(* IEC 61131-3 sources: SortJet_MasterSPS_Aufbau.fbsproj/08_POUs/Basis Funktionen, 41 files *)

(* ---- AuftragsdatenPruefen.fn.st ---- *)
(* METADATA
{
	"v3Meta": {
		"objectGuid": "657d7773-50f6-4a46-b86f-6fc5131c38e4"
	}
}
*)
FUNCTION AuftragsdatenPruefen : BOOL
VAR_INPUT

  // WORD
  wpMmiNummer  : WORD; // Stationsnummer von der die Auftraege geprueft werden sollen
  wpWandNr     : WORD; // Wandnummer von der die Auftraege geprueft werden sollen

  // STRUKT
  pData   : Auftragsdaten_ST;

END_VAR
VAR
  Basis : REFERENCE TO StationBasisParameter_ST;
END_VAR
Basis REF= getBasis(wpMmiNummer);
AuftragsdatenPruefen := TRUE;

// Glaslänge
IF ( pData.rAuftragsLaenge > Basis.stMKs.stGlasdaten[wpWandNr].rlMaxGlasLaenge ) THEN
  wpgFehlerdaten[0] := wpMmiNummer;
  wpgFehlerdaten[1] := REAL_TO_WORD(Basis.stMKs.stGlasdaten[wpWandNr].rlMaxGlasLaenge);
  wpgFehlerdaten[2] := REAL_TO_WORD(pData.rAuftragsLaenge);
  SpsError( eFehler_Station,
            cMELDUNG_AUFTRAGSDATEN_GLAS_ZU_LANG,
            wpMmiNummer,
            AutomatikkreisBestimmen(wpMmiNummer),
            wpgFehlerdaten );
  AuftragsdatenPruefen:=FALSE;
END_IF

IF ( pData.rAuftragsLaenge < Basis.stMKs.stGlasdaten[wpWandNr].rlMinGlasLaenge ) THEN
  wpgFehlerdaten[0] := wpMmiNummer;
  wpgFehlerdaten[1] := REAL_TO_WORD(Basis.stMKs.stGlasdaten[wpWandNr].rlMinGlasLaenge);
  wpgFehlerdaten[2] := REAL_TO_WORD(pData.rAuftragsLaenge);
  SpsError( eFehler_Station,
            cMELDUNG_AUFTRAGSDATEN_GLAS_ZU_KURZ,
            wpMmiNummer,
            AutomatikkreisBestimmen(wpMmiNummer),
            wpgFehlerdaten );
  AuftragsdatenPruefen:=FALSE;
END_IF

// Glashöhe
IF ( pData.rAuftragsHoehe > Basis.stMKs.stGlasdaten[wpWandNr].rlMaxGlasHoehe ) THEN
  wpgFehlerdaten[0] := wpMmiNummer;
  wpgFehlerdaten[1] := REAL_TO_WORD(Basis.stMKs.stGlasdaten[wpWandNr].rlMaxGlasHoehe);
  wpgFehlerdaten[2] := REAL_TO_WORD(pData.rAuftragsHoehe);
  SpsError( eFehler_Station,
            cMELDUNG_AUFTRAGSDATEN_GLAS_ZU_HOCH,
            wpMmiNummer,
            AutomatikkreisBestimmen(wpMmiNummer),
            wpgFehlerdaten );
  AuftragsdatenPruefen:=FALSE;
END_IF

IF ( pData.rAuftragsHoehe <  Basis.stMKs.stGlasdaten[wpWandNr].rlMinGlasHoehe ) THEN
  wpgFehlerdaten[0] := wpMmiNummer;
  wpgFehlerdaten[1] := REAL_TO_WORD(Basis.stMKs.stGlasdaten[wpWandNr].rlMinGlasHoehe);
  wpgFehlerdaten[2] := REAL_TO_WORD(pData.rAuftragsHoehe);
  SpsError( eFehler_Station,
            cMELDUNG_AUFTRAGSDATEN_GLAS_ZU_NIEDRIG,
            wpMmiNummer,
            AutomatikkreisBestimmen(wpMmiNummer),
            wpgFehlerdaten );
  AuftragsdatenPruefen:=FALSE;
END_IF

// Glasdicke
IF ( pData.rAuftragsDicke > Basis.stMKs.stGlasdaten[wpWandNr].rlMaxGlasDicke ) THEN
  wpgFehlerdaten[0] := wpMmiNummer;
  wpgFehlerdaten[1] := REAL_TO_WORD(Basis.stMKs.stGlasdaten[wpWandNr].rlMaxGlasDicke);
  wpgFehlerdaten[2] := REAL_TO_WORD(pData.rAuftragsDicke);
  SpsError( eFehler_Station,
            cMELDUNG_AUFTRAGSDATEN_GLAS_ZU_DICK,
            wpMmiNummer,
            AutomatikkreisBestimmen(wpMmiNummer),
            wpgFehlerdaten );
  AuftragsdatenPruefen := FALSE;
END_IF

IF ( pData.rAuftragsDicke < Basis.stMKs.stGlasdaten[wpWandNr].rlMinGlasDicke ) THEN
  wpgFehlerdaten[0] := wpMmiNummer;
  wpgFehlerdaten[1] := REAL_TO_WORD(Basis.stMKs.stGlasdaten[wpWandNr].rlMinGlasDicke);
  wpgFehlerdaten[2] := REAL_TO_WORD(pData.rAuftragsDicke);
  SpsError( eFehler_Station,
            cMELDUNG_AUFTRAGSDATEN_GLAS_ZU_DUENN,
            wpMmiNummer,
            AutomatikkreisBestimmen(wpMmiNummer),
            wpgFehlerdaten );
  AuftragsdatenPruefen := FALSE;
END_IF
END_FUNCTION

(* ---- AuftragsdatenUmkopieren.fn.st ---- *)
(* METADATA
{
	"v3Meta": {
		"objectGuid": "c0c5d446-5c0c-4964-91ed-f4edd34c4197"
	}
}
*)
FUNCTION AuftragsdatenUmkopieren : Auftragsdaten_ST
VAR_INPUT

  // BOOL
  bpAuswahlTransferstation_2  : BOOL := FALSE;
  bpAnwahlDurchtransport : BOOL := FALSE;

  // STRUCT
  stpAuftrag : Auftragsdaten_ST;

END_VAR
VAR

  // STRUCT
  stMerkerAuftrag  : Auftragsdaten_ST;

END_VAR
//-------------------------------------------------------------------------------------------------
// BAUSTEIN: LOGIK
//-------------------------------------------------------------------------------------------------

(* Hinweis:
   - Auftrag zwischenspeichern
*)
stMerkerAuftrag := stpAuftrag;

(* Hinweis:
   - Auftrag manipulieren
*)
IF ( NOT bpAuswahlTransferstation_2 AND NOT bpAnwahlDurchtransport ) THEN

  stMerkerAuftrag.wStationsNr            := stpAuftrag.wTransferstationsNr1;
  stMerkerAuftrag.wStationsWand          := stpAuftrag.wTransferwand;
  stMerkerAuftrag.rStationsZielposition  := stpAuftrag.rTransferposition1;
  stMerkerAuftrag.rVorabPosition         := stpAuftrag.rTransferposition1;

  stMerkerAuftrag.wTransferstationsNr1   := stpAuftrag.wStationsNr;
  stMerkerAuftrag.rTransferposition1     := stpAuftrag.rStationsZielposition;
  stMerkerAuftrag.wTransferwand          := stpAuftrag.wStationsWand;

ELSIF ( bpAnwahlDurchtransport ) THEN

  stMerkerAuftrag.wStationsNr            := stpAuftrag.wTransferstationsNr2;
  stMerkerAuftrag.wStationsWand          := stpAuftrag.wTransferwand;
  stMerkerAuftrag.rStationsZielposition  := stpAuftrag.rTransferposition2;
  stMerkerAuftrag.rVorabPosition         := stpAuftrag.rTransferposition2;

  stMerkerAuftrag.wTransferstationsNr2   := stpAuftrag.wStationsNr;
  stMerkerAuftrag.rTransferposition2     := stpAuftrag.rStationsZielposition;
  stMerkerAuftrag.wTransferwand          := stpAuftrag.wStationsWand;

ELSE
  stMerkerAuftrag.wStationsNr            := stpAuftrag.wTransferstationsNr2;
  stMerkerAuftrag.wStationsWand          := stpAuftrag.wTransferwand;
  stMerkerAuftrag.rStationsZielposition  := stpAuftrag.rTransferposition2;
  stMerkerAuftrag.rVorabPosition         := stpAuftrag.rTransferposition2;

  stMerkerAuftrag.wTransferstationsNr1   := stpAuftrag.wStationsNr;
  stMerkerAuftrag.rTransferposition1     := stpAuftrag.rStationsZielposition;
  stMerkerAuftrag.wTransferwand          := stpAuftrag.wStationsWand;

END_IF

AuftragsdatenUmkopieren := stMerkerAuftrag;
END_FUNCTION

(* ---- AutomatikAktiv.fn.st ---- *)
(* METADATA
{
	"v3Meta": {
		"objectGuid": "339b2ef9-3f23-482c-98f4-06c495d9a955"
	}
}
*)
FUNCTION AutomatikAktiv : BOOL
VAR_INPUT
  wpMmiNummer : WORD;
END_VAR
VAR
  wlIndex : WORD;
  Basis   : REFERENCE TO StationBasisParameter_ST;
END_VAR

// Hinweis:
// - Prueft ob einer der Automatikkreise der Station (Shuttle, TS, Station, Faecherwagen, Fremdanlage) aktiv ist
// - Die Basis wird ueber getBasis bestimmt
// - Unbekannte Nummer oder nicht zugewiesene MK => FALSE
// - Ein nicht belegter Automatikkreis (0) beendet die Pruefung
AutomatikAktiv := FALSE;

Basis REF= getBasis( wpMmiNummer );

IF NOT __ISVALIDREF( Basis ) THEN
  RETURN;
END_IF

IF NOT __ISVALIDREF( Basis.stMKs ) THEN
  RETURN;
END_IF

FOR wlIndex := cERSTER_AUTOMATIKKREIS TO cANZAHL_AUTOMATIKKREISE DO

  IF Basis.stMKs.eaAutomatikkreis[wlIndex] = 0 THEN
    RETURN;
  END_IF

  IF M_Automatik_Aktiv[Basis.stMKs.eaAutomatikkreis[wlIndex]] THEN
    AutomatikAktiv := TRUE;
    RETURN;
  END_IF

END_FOR
END_FUNCTION

(* ---- AutomatikFehlerSetzen.fn.st ---- *)
(* METADATA
{
	"v3Meta": {
		"objectGuid": "10c1b2d6-77ce-44d1-9dc1-390f3ff85d9b"
	}
}
*)
FUNCTION AutomatikFehlerSetzen : BOOL
VAR_INPUT
  eaAutomatikkreise : ARRAY[cERSTER_AUTOMATIKKREIS..cANZAHL_AUTOMATIKKREISE] OF Automatikkreis_EN;
  abpFehler : REFERENCE TO ARRAY[cERSTER_AUTOMATIKKREIS..cLETZTER_AUTOMATIKKREIS] OF BOOL;
END_VAR
VAR
  wlIndex: WORD;
END_VAR

FOR wlIndex := cERSTER_AUTOMATIKKREIS TO cANZAHL_AUTOMATIKKREISE DO

  IF eaAutomatikkreise[wlIndex] <> 0 THEN
    abpFehler[eaAutomatikkreise[wlIndex]] := TRUE;
  END_IF

END_FOR

AutomatikFehlerSetzen := TRUE;
END_FUNCTION

(* ---- AutomatikFehlerTransfershuttleSetzen.fn.st ---- *)
(* METADATA
{
	"v3Meta": {
		"objectGuid": "9a4c379e-af86-4c9e-b628-bbb819ee7aed"
	}
}
*)
FUNCTION AutomatikFehlerTransfershuttleSetzen : BOOL
VAR_INPUT
  eaAutomatikkreise    : ARRAY[cERSTER_AUTOMATIKKREIS..cANZAHL_AUTOMATIKKREISE] OF Automatikkreis_EN;
  abpFehler            : REFERENCE TO ARRAY[cERSTER_AUTOMATIKKREIS..cLETZTER_AUTOMATIKKREIS] OF BOOL;
  wSpeicherseiteFehler : BYTE; // cSPEICHER_EINLAUFSEITE oder cSPEICHER_AUSLAUFSEITE
END_VAR

// Hinweis:
// - Ein TS liegt meist als Trennglied unter dem Speicher in 2 AKs:
//   AK 1 = Einlaufseite, AK 2 = Auslaufseite
// - Welche Seite betroffen ist (Ein-/Austransport, rueckwaerts, Betriebsstopp)
//   entscheidet der Aufrufer in Job_Shuttle

// TS hat nur einen AK
IF ( eaAutomatikkreise[1] <> 0 AND eaAutomatikkreise[2] = 0 ) THEN
  abpFehler[eaAutomatikkreise[1]] := TRUE;

// TS hat 2 AK
ELSIF ( eaAutomatikkreise[1] <> 0 AND eaAutomatikkreise[2] <> 0 ) THEN
  IF ( wSpeicherseiteFehler = cSPEICHER_EINLAUFSEITE ) THEN
    abpFehler[eaAutomatikkreise[1]] := TRUE;
  ELSIF ( wSpeicherseiteFehler = cSPEICHER_AUSLAUFSEITE ) THEN
    abpFehler[eaAutomatikkreise[2]] := TRUE;
  END_IF
END_IF

AutomatikFehlerTransfershuttleSetzen := TRUE;
END_FUNCTION

(* ---- AutomatikkreisBestimmen.fn.st ---- *)
(* METADATA
{
	"v3Meta": {
		"objectGuid": "9ed7362d-6e8b-45fc-aaf5-a3cbb726335b"
	}
}
*)
FUNCTION AutomatikkreisBestimmen : Automatikkreis_EN
VAR_INPUT
  wpMmiNummer : WORD;
END_VAR
VAR
  Basis : REFERENCE TO StationBasisParameter_ST;
END_VAR

// Hinweis:
// - Erster Automatikkreis der Station (Shuttle, TS, Station, Faecherwagen, Fremdanlage) ueber getBasis
// - Unbekannte Nummer oder nicht zugewiesene MK => 0
AutomatikkreisBestimmen := 0;

Basis REF= getBasis( wpMmiNummer );

IF NOT __ISVALIDREF( Basis ) THEN
  RETURN;
END_IF

IF NOT __ISVALIDREF( Basis.stMKs ) THEN
  RETURN;
END_IF

AutomatikkreisBestimmen := Basis.stMKs.eaAutomatikkreis[cERSTER_AUTOMATIKKREIS];
END_FUNCTION

(* ---- BitToggleWord.fn.st ---- *)
(* METADATA
{
	"v3Meta": {
		"objectGuid": "aa0bc2f8-efb2-48a1-91f1-3637f8b86daf"
	}
}
*)
FUNCTION BitToggleWord : WORD
VAR_INPUT

  // WORD
  IN : WORD;

  // INT
  POS : INT;

END_VAR
//-------------------------------------------------------------------------------------------------
// BAUSTEIN: LOGIK
//-------------------------------------------------------------------------------------------------

(* Hinweis:
   - Diese Funktion setzt in einem WORD ein BIT an einer Position
     => Oscat-Lib
*)
BitToggleWord := SHL(WORD#1, POS) XOR IN;
END_FUNCTION

(* ---- checkSafetyCircuitAffectsComponent.fn.st ---- *)
(* METADATA
{
	"v3Meta": {
		"objectGuid": "b2891e00-4397-4c85-8733-7380e4011fc3"
	}
}
*)
FUNCTION checkSafetyCircuitAffectsComponent : BOOL
VAR_INPUT
  StationData  : REFERENCE TO StationBasisParameter_ST;
  SaftyCircuit : WORD;              // Sicherheitskreis
  eKomponente  : SK_Komponente_EN;  // Abgefragte Komponente (eSKKomponente_Alles = jeder SK zaehlt)
END_VAR
VAR
  wIndexMK : WORD := 0;
END_VAR
// Prueft, ob ein Sicherheitskreis die angegebene Komponente der Station abschaltet.
// - eSKKomponente_Alles: jeder SK der Station zaehlt -> TRUE
// - Standard (keine Teilabschaltung fuer diesen SK konfiguriert): SK schaltet alles ab -> TRUE
// - Mit Teilabschaltung: SK schaltet nur die markierten Komponenten ab

checkSafetyCircuitAffectsComponent := TRUE;

IF ( eKomponente = eSKKomponente_Alles ) THEN
  RETURN;
END_IF

FOR wIndexMK := 0 TO cANZAHL_SICHERHEITSKREISE DO
  IF     ( StationData.stMKs.astSicherheitskreisTeilabschaltung[wIndexMK].eSicherheitskreis = SaftyCircuit )
     AND StationData.stMKs.astSicherheitskreisTeilabschaltung[wIndexMK].bTeilabschaltung
  THEN
    CASE eKomponente OF
      eSKKomponente_Glastransport:   checkSafetyCircuitAffectsComponent := StationData.stMKs.astSicherheitskreisTeilabschaltung[wIndexMK].bGlastransport;
      eSKKomponente_Geblaese:        checkSafetyCircuitAffectsComponent := StationData.stMKs.astSicherheitskreisTeilabschaltung[wIndexMK].bGeblaese;
      eSKKomponente_Drehen:          checkSafetyCircuitAffectsComponent := StationData.stMKs.astSicherheitskreisTeilabschaltung[wIndexMK].bDrehen;
      eSKKomponente_Kippen:          checkSafetyCircuitAffectsComponent := StationData.stMKs.astSicherheitskreisTeilabschaltung[wIndexMK].bKippen;
      eSKKomponente_Querfahrt:       checkSafetyCircuitAffectsComponent := StationData.stMKs.astSicherheitskreisTeilabschaltung[wIndexMK].bQuerfahrt;
      eSKKomponente_Pneumatik:       checkSafetyCircuitAffectsComponent := StationData.stMKs.astSicherheitskreisTeilabschaltung[wIndexMK].bPneumatik;
      eSKKomponente_Greifer:         checkSafetyCircuitAffectsComponent := StationData.stMKs.astSicherheitskreisTeilabschaltung[wIndexMK].bGreifer;
      eSKKomponente_Wandverstellung: checkSafetyCircuitAffectsComponent := StationData.stMKs.astSicherheitskreisTeilabschaltung[wIndexMK].bWandverstellung;
      eSKKomponente_Messachse:       checkSafetyCircuitAffectsComponent := StationData.stMKs.astSicherheitskreisTeilabschaltung[wIndexMK].bMessachse;
    END_CASE
    RETURN;
  END_IF
END_FOR
END_FUNCTION

(* ---- checkSafetyCircuits.fn.st ---- *)
(* METADATA
{
	"v3Meta": {
		"objectGuid": "a5602391-f145-45a7-88a7-cf2977d4c874"
	}
}
*)
FUNCTION checkSafetyCircuits : BOOL
VAR_INPUT
  StationData  : REFERENCE TO StationBasisParameter_ST;
  SaftyCircuit : WORD;
END_VAR
VAR
  wIndexMK : WORD := 0;
END_VAR
// It will checked if the safety circuit configured for this station

checkSafetyCircuits := FALSE;

FOR wIndexMK := 0 TO cANZAHL_SICHERHEITSKREISE DO
  IF ( SaftyCircuit = StationData.stMKs.eaSicherheitskreis[wIndexMK] ) THEN
    checkSafetyCircuits := TRUE;
    EXIT;
  END_IF
END_FOR
END_FUNCTION

(* ---- checkSafetyCircuitsClosed.fn.st ---- *)
(* METADATA
{
	"v3Meta": {
		"objectGuid": "1a45708a-46ce-48f5-a3b2-b0c20261c8e1"
	}
}
*)
FUNCTION checkSafetyCircuitsClosed : BOOL
VAR_INPUT
  StationData : REFERENCE TO StationBasisParameter_ST;
  eKomponente : SK_Komponente_EN := eSKKomponente_Alles; // Optional: Pruefung fuer eine Komponente (beruecksichtigt Teilabschaltung), Standard: jeder SK zaehlt
END_VAR
VAR
  arrCircuits : ARRAY[cERSTER_SICHERHEITSKREIS..cLETZTER_SICHERHEITSKREIS] OF BOOL;
  wIndex   : WORD := 0;
  wIndexMK : WORD := 0;
END_VAR
// It will checked if the safety circuit is activ

checkSafetyCircuitsClosed := TRUE;

FOR wIndex := cERSTER_SICHERHEITSKREIS TO cLETZTER_SICHERHEITSKREIS DO
  arrCircuits[wIndex] := Sicherheitskreis[wIndex].bpSicherheitskreisGeschlossen;
END_FOR

FOR wIndex := cERSTER_SICHERHEITSKREIS TO cLETZTER_SICHERHEITSKREIS DO
  FOR wIndexMK := 0 TO cANZAHL_SICHERHEITSKREISE DO
    IF ( wIndex = StationData.stMKs.eaSicherheitskreis[wIndexMK] ) THEN
      IF NOT arrCircuits[wIndex] AND checkSafetyCircuitAffectsComponent(StationData, wIndex, eKomponente) THEN
        checkSafetyCircuitsClosed := FALSE;
      END_IF
    END_IF
  END_FOR
END_FOR
END_FUNCTION

(* ---- checkSafetyCircuitsClosedFromAutomaticCircuit.fn.st ---- *)
(* METADATA
{
	"v3Meta": {
		"objectGuid": "6a4b769b-603d-4996-8e76-e26c1b994362"
	}
}
*)
FUNCTION checkSafetyCircuitsClosedFromAutomaticCircuit : BOOL
VAR_INPUT

  // WORD
  wlAutomatikkreis : WORD;

  // BOOL
  bNurStartBlockierende : BOOL := FALSE; // TRUE: nur Sicherheitskreise beruecksichtigen, die Systemcheck und Initialisierung blockieren [MK bBlockiertStart]

END_VAR
VAR
  // BOOL
  findInWORDArray               : BOOL;
  bSicherheitskreisIstDurchgang : BOOL;

  // WORD
  wlIndexSicherheitskreis : WORD;

  // ENUM
  INDEX : Automatikkreis_EN;

END_VAR

// DIESE FUNKTION BERÜCKSICHTIGT KEINE DURCHGÄNGE !!!
checkSafetyCircuitsClosedFromAutomaticCircuit := TRUE;

FOR wlIndexSicherheitskreis := cERSTER_SICHERHEITSKREIS TO cLETZTER_SICHERHEITSKREIS DO

  bSicherheitskreisIstDurchgang := FALSE;

  FOR INDEX := cERSTER_DURCHGANG TO cANZAHL_DURCHGANGE DO
    IF apgMKDurchgang[INDEX].eZuBlockierenderSK = wlIndexSicherheitskreis THEN
      bSicherheitskreisIstDurchgang := TRUE;
      EXIT;
    END_IF
  END_FOR

  IF NOT bSicherheitskreisIstDurchgang THEN

    findInWORDArray := FALSE;

    FOR INDEX := cERSTER_AUTOMATIKKREIS TO cLETZTER_AUTOMATIKKREIS DO
      IF apgMKSicherheiskreis[wlIndexSicherheitskreis].eaAutomatikkreis[INDEX] = wlAutomatikkreis THEN
        findInWORDArray := TRUE;
        EXIT;
      END_IF
    END_FOR

    IF findInWORDArray AND ( NOT bNurStartBlockierende OR apgMKSicherheiskreis[wlIndexSicherheitskreis].bBlockiertStart ) THEN
      checkSafetyCircuitsClosedFromAutomaticCircuit :=
                                                      checkSafetyCircuitsClosedFromAutomaticCircuit
                                                      AND Sicherheitskreis[wlIndexSicherheitskreis].bpSicherheitskreisGeschlossen;
    END_IF

  END_IF

END_FOR
END_FUNCTION

(* ---- checkSafetyCircuitsConfigured.fn.st ---- *)
(* METADATA
{
	"v3Meta": {
		"objectGuid": "dcded4cc-d766-4c84-a212-2fe6cc93f6db"
	}
}
*)
FUNCTION checkSafetyCircuitsConfigured : BOOL
VAR_INPUT
  StationData : REFERENCE TO StationBasisParameter_ST;
END_VAR
VAR
  wIndexMK : WORD := 0;
END_VAR

// It will checked if a safety circuit is configured

checkSafetyCircuitsConfigured := FALSE;

IF NOT __ISVALIDREF(StationData.stMKs) OR_ELSE StationData.stMKs.bDeaktivieren THEN
  RETURN;
END_IF

FOR wIndexMK := 0 TO cANZAHL_SICHERHEITSKREISE DO
  IF ( StationData.stMKs.eaSicherheitskreis[wIndexMK] <> eSicherheitskreis_Undefiniert ) THEN
    checkSafetyCircuitsConfigured := TRUE;
    EXIT;
  END_IF
END_FOR
END_FUNCTION

(* ---- checkSafetyCircuitsNotBlocked.fn.st ---- *)
(* METADATA
{
	"v3Meta": {
		"objectGuid": "93537a12-23ea-4a31-94f7-53154eb0b75f"
	}
}
*)
FUNCTION checkSafetyCircuitsNotBlocked : BOOL
VAR_INPUT
  StationData : REFERENCE TO StationBasisParameter_ST;
  eKomponente : SK_Komponente_EN := eSKKomponente_Alles; // Optional: Pruefung fuer eine Komponente (beruecksichtigt Teilabschaltung), Standard: jeder SK zaehlt
END_VAR
VAR
  arrCircuits : ARRAY[cERSTER_SICHERHEITSKREIS..cLETZTER_SICHERHEITSKREIS] OF BOOL;
  wIndex   : WORD := 0;
  wIndexMK : WORD := 0;
END_VAR
// It will checked if the safety circuit is activ

checkSafetyCircuitsNotBlocked := TRUE;

FOR wIndex := cERSTER_SICHERHEITSKREIS TO cLETZTER_SICHERHEITSKREIS DO
  arrCircuits[wIndex] :=         Sicherheitskreis[wIndex].bpSicherheitskreisGeschlossen
                                 AND NOT Sicherheitskreis[wIndex].bpStationenBlocken
                                 AND NOT Sicherheitskreis[wIndex].bpAnforderungSKGestellt
                                 AND NOT Sicherheitskreis[wIndex].bpAnforderungSicherheitkreisAusloesen;
END_FOR

FOR wIndex := cERSTER_SICHERHEITSKREIS TO cLETZTER_SICHERHEITSKREIS DO
  FOR wIndexMK := 0 TO cANZAHL_SICHERHEITSKREISE DO
    IF ( wIndex = StationData.stMKs.eaSicherheitskreis[wIndexMK] ) THEN
      IF ( ( NOT arrCircuits[wIndex] ) AND ( NOT bgSicherheitstechnikBruecken ) AND checkSafetyCircuitAffectsComponent(StationData, wIndex, eKomponente) ) THEN
        checkSafetyCircuitsNotBlocked := FALSE;
        EXIT;
      END_IF
    END_IF
  END_FOR
END_FOR
END_FUNCTION

(* ---- checkSafetyCircuitsRequested.fn.st ---- *)
(* METADATA
{
	"v3Meta": {
		"objectGuid": "c6e29fd6-ba36-47ef-8c35-03485548b8fc"
	}
}
*)
FUNCTION checkSafetyCircuitsRequested : BOOL
VAR_INPUT
  StationData : REFERENCE TO StationBasisParameter_ST;
  eKomponente : SK_Komponente_EN := eSKKomponente_Alles; // Optional: Pruefung fuer eine Komponente (beruecksichtigt Teilabschaltung), Standard: jeder SK zaehlt
END_VAR
VAR
  arrCircuits : ARRAY[cERSTER_SICHERHEITSKREIS..cLETZTER_SICHERHEITSKREIS] OF BOOL;
  wIndex   : WORD := 0;
  wIndexMK : WORD := 0;
END_VAR
// It will checked if the safety circuit is requested

checkSafetyCircuitsRequested := TRUE;

FOR wIndex := cERSTER_SICHERHEITSKREIS TO cLETZTER_SICHERHEITSKREIS DO
  arrCircuits[wIndex] :=         Sicherheitskreis[wIndex].bpSicherheitskreisGeschlossen
                                 AND NOT Sicherheitskreis[wIndex].bpAnforderungSKGestellt;
END_FOR

FOR wIndex := cERSTER_SICHERHEITSKREIS TO cLETZTER_SICHERHEITSKREIS DO

  FOR wIndexMK := 0 TO cANZAHL_SICHERHEITSKREISE DO
    IF ( wIndex = StationData.stMKs.eaSicherheitskreis[wIndexMK] ) THEN
      IF NOT arrCircuits[wIndex] AND checkSafetyCircuitAffectsComponent(StationData, wIndex, eKomponente) THEN
        checkSafetyCircuitsRequested := FALSE;
      END_IF
    END_IF
  END_FOR
END_FOR
END_FUNCTION

(* ---- DEC.fn.st ---- *)
(* METADATA
{
	"v3Meta": {
		"objectGuid": "e4081493-5d9a-4e63-8c4b-cba513ba3d02"
	}
}
*)
{attribute 'excludefrombuild'}
FUNCTION DEC : INT
VAR_INPUT
  iWert    : INT;
  iMinuend : INT;
END_VAR

(* Hinweis:
   - Funktion zum reduzieren der Eingangsvariablen X um 1.
*)
DEC := iWert - iMinuend;
END_FUNCTION

(* ---- findInWORDArray.fn.st ---- *)
(* METADATA
{
	"v3Meta": {
		"objectGuid": "27266190-4c13-454c-9114-87648310c4ec"
	}
}
*)
FUNCTION findInWORDArray : BOOL
VAR_INPUT
  awpArray : ARRAY[1..10] OF WORD;
  wpValueToFind : WORD;
END_VAR
VAR
  INDEX : WORD;
END_VAR

findInWORDArray := FALSE;

FOR INDEX := 1 TO 10 DO

  IF awpArray[INDEX] = wpValueToFind THEN
    findInWORDArray := TRUE;
    EXIT;
  END_IF

END_FOR
END_FUNCTION

(* ---- getAnzahlSystemcheckZyklen.fn.st ---- *)
(* METADATA
{
	"v3Meta": {
		"objectGuid": "64956d77-da35-4a2e-90f0-c969659e6e9b"
	}
}
*)
FUNCTION getAnzahlSystemcheckZyklen : WORD
VAR_INPUT
END_VAR
VAR
  wIndex : WORD;
  bByte  : BYTE;
  ptNull : REFERENCE TO BYTE := 0;
END_VAR

getAnzahlSystemcheckZyklen := 0;

// Alle Shuttles durchlaufen
FOR wIndex := cERSTES_SHUTTLE TO cLETZTES_SHUTTLE DO
  // Null-Pointer wenn kein Zyklus in den MKs zugewiesen wurde
  IF starrShuttleBasisParameter[wIndex].stMKs.eSystemcheckZyklus = eSystemcheckZyklus_Undefiniert THEN
    SysExceptGenerateException( RtsExceptions.RTSEXCPT_ARRAYBOUNDS );
  //bByte := ptNull; (*cause access violation *)
  ELSE // Ansonsten den definierten Zyklus in das Array übernehmen
    // Neuer höherer Wert? Dann wegspeichern
    IF getAnzahlSystemcheckZyklen < starrShuttleBasisParameter[wIndex].stMKs.eSystemcheckZyklus THEN
      getAnzahlSystemcheckZyklen := starrShuttleBasisParameter[wIndex].stMKs.eSystemcheckZyklus;
    END_IF
  END_IF
END_FOR

// Alle Stationen durchlaufen
FOR wIndex := cERSTE_STATION TO cLETZTE_STATION DO
  // Null-Pointer wenn kein Zyklus in den MKs zugewiesen wurde
  IF NOT __ISVALIDREF(starrStationBasisParameter[wIndex].stMKs) THEN
    CONTINUE;
  ELSIF starrStationBasisParameter[wIndex].stMKs.eSystemcheckZyklus = eSystemcheckZyklus_Undefiniert AND NOT starrStationBasisParameter[wIndex].stMKs.bDeaktivieren THEN
    SysExceptGenerateException( RtsExceptions.RTSEXCPT_ARRAYBOUNDS );
  //bByte := ptNull; (*cause access violation *)
  ELSE // Ansonsten den definierten Zyklus in das Array übernehmen
    // Neuer höherer Wert? Dann wegspeichern
    IF getAnzahlSystemcheckZyklen < starrStationBasisParameter[wIndex].stMKs.eSystemcheckZyklus THEN
      getAnzahlSystemcheckZyklen := starrStationBasisParameter[wIndex].stMKs.eSystemcheckZyklus;
    END_IF
  END_IF
END_FOR

// Null-Pointer wenn kein Ergebnis gefunden wurde (fehlerhafter Zustand)
IF ( getAnzahlSystemcheckZyklen = 0 ) THEN
  SysExceptGenerateException( RtsExceptions.RTSEXCPT_ARRAYBOUNDS );
//bByte := ptNull; (*cause access violation *)
END_IF
END_FUNCTION

(* ---- getAuftragsdaten.fn.st ---- *)
(* METADATA
{
	"v3Meta": {
		"objectGuid": "e09c3e56-23fc-432f-9a18-960dccfa6275"
	}
}
*)
FUNCTION getAuftragsdaten : REFERENCE TO Auftragsdaten_ST
VAR_INPUT

  // WORD
  wpMmiNummer  : WORD; // Stationsnummer, deren aktueller Auftrag geliefert werden soll
  wpWand       : WORD; // Wand (nur Shuttles und Stationen)

END_VAR
// Hinweis:
// - Gegenstueck zu getBasis: liefert den aktuellen Job-Auftrag einer Station
// - Ungueltige Nummer oder Wand => ungueltige Referenz (Aufrufer prueft mit __ISVALIDREF)
CASE wpMmiNummer OF

  cERSTES_SHUTTLE..cLETZTES_SHUTTLE:
    IF ( PruefungWertImIntervall( wpWand, cWAND_1, cANZAHL_WAENDE ) ) THEN
      getAuftragsdaten REF= Job_Shuttle.AuftragsdatenWand[wpMmiNummer, wpWand];
    END_IF

  cERSTES_TRANSFERSHUTTLE..cLETZTES_TRANSFERSHUTTLE:
    getAuftragsdaten REF= Job_Shuttle.AuftragsdatenTransfershuttle[wpMmiNummer];

  cERSTE_STATION..cLETZTE_STATION:
    IF ( PruefungWertImIntervall( wpWand, cWAND_1, cANZAHL_WAENDE ) ) THEN
      getAuftragsdaten REF= Job_Stationen.AuftragsdatenWand[wpMmiNummer, wpWand];
    END_IF

  cERSTE_FREMDANLAGE_AUSLAUF..cLETZTE_FREMDANLAGE_EINLAUF:
    getAuftragsdaten REF= Job_Fremdanlage.AuftragsdatenFremdanlage[wpMmiNummer];

END_CASE
END_FUNCTION

(* ---- getBasis.fn.st ---- *)
(* METADATA
{
	"v3Meta": {
		"objectGuid": "cb0abf05-d74d-4b59-9143-e94abaf551fa"
	}
}
*)
FUNCTION getBasis : REFERENCE TO  StationBasisParameter_ST
VAR_INPUT

  // WORD
  wpMmiNummer  : WORD; // Stationsnummer von der die Auftraege geprueft werden sollen

END_VAR
CASE wpMmiNummer OF

  cERSTES_SHUTTLE..cLETZTES_SHUTTLE:
    getBasis REF= starrShuttleBasisParameter[wpMmiNummer];

  cERSTES_TRANSFERSHUTTLE..cLETZTES_TRANSFERSHUTTLE:
    getBasis REF= starrTransfershuttleBasisParameter[wpMmiNummer];

  cERSTE_STATION..cLETZTE_STATION:
    getBasis REF= starrStationBasisParameter[wpMmiNummer];

  cERSTE_FAECHERWAGENSTATIONS_NR..cLETZTE_FAECHERWAGENSTATIONS_NR:
    getBasis REF= starrFaecherwagenBasisParameter[wpMmiNummer];

  cERSTE_FREMDANLAGE_EINLAUF..cLETZTE_FREMDANLAGE_EINLAUF:
    getBasis REF= starrFremdanlageEinlaufStationBasisParameter[wpMmiNummer];

  cERSTE_FREMDANLAGE_AUSLAUF..cLETZTE_FREMDANLAGE_AUSLAUF:
    getBasis REF= starrFremdanlageAuslaufStationBasisParameter[wpMmiNummer];

END_CASE
END_FUNCTION

(* ---- GetBitFromWord.fn.st ---- *)
(* METADATA
{
	"v3Meta": {
		"objectGuid": "4ac38ee7-2639-4587-9c58-5882c3701cd8"
	}
}
*)
FUNCTION GetBitFromWord : Bool
VAR_INPUT
  Value : WORD;   // Das Wort, aus dem du die Bits auslesen willst
  Index : Word;    // Welches Bit (0..15)
END_VAR
VAR
END_VAR

GetBitFromWord := (Value AND SHL(1, Index)) <> 0;
END_FUNCTION

(* ---- getRealShuttleMaxPos.fn.st ---- *)
(* METADATA
{
	"v3Meta": {
		"objectGuid": "fdbd0502-3da4-4780-aa1a-b043617e0f01"
	}
}
*)
FUNCTION getRealShuttleMaxPos : REAL
VAR_INPUT
  wShuttleNummer : WORD;
END_VAR

getRealShuttleMaxPos := aShuttle[wShuttleNummer].Querfahrt.Antrieb.rpMaxPosition;
END_FUNCTION

(* ---- getRealShuttleMinPos.fn.st ---- *)
(* METADATA
{
	"v3Meta": {
		"objectGuid": "77446a83-5414-4511-a85e-8d0f27ae2e7b"
	}
}
*)
FUNCTION getRealShuttleMinPos : REAL
VAR_INPUT
  wShuttleNummer : WORD;
END_VAR

getRealShuttleMinPos := aShuttle[wShuttleNummer].Querfahrt.Antrieb.rpMinPosition;
END_FUNCTION

(* ---- GlasGewichtErmitteln.fn.st ---- *)
(* METADATA
{
	"v3Meta": {
		"objectGuid": "bd924e48-93d5-4f05-bff1-59051efc4e7c"
	}
}
*)
FUNCTION GlasGewichtErmitteln : REAL
VAR_INPUT

  // REAL
  rpGlaslaenge  : REAL := REAL#0; // [mm] -> Wert in mm
  rpGlasbreite  : REAL := REAL#0; // [mm] -> Wert in mm
  rpGlasstaerke : REAL := REAL#0; // [mm] -> Wert in mm

END_VAR
VAR

  // REAL
  rlErgebnis : REAL := REAL#0;
  rlLaenge   : REAL := REAL#0; // [mm] -> Wert in dm [UMRECHNUNG]
  rlBreite   : REAL := REAL#0; // [mm] -> Wert in dm [UMRECHNUNG]
  rlStaerke  : REAL := REAL#0; // [mm] -> Wert in dm [UMRECHNUNG]

END_VAR

VAR CONSTANT

  // WORD
  cUMRECHNUNG_MM_IN_DM      : REAL := 100.0;

  // REAL
  cSPEZIFISCHES_GLASGEWICHT : REAL := REAL#2.5; //IN kg/dm³

END_VAR

rlErgebnis := REAL#0;

rlLaenge  := rpGlaslaenge / cUMRECHNUNG_MM_IN_DM;
rlBreite  := rpGlasbreite / cUMRECHNUNG_MM_IN_DM;
rlStaerke := rpGlasstaerke/ cUMRECHNUNG_MM_IN_DM;

GlasGewichtErmitteln := ( ( rlLaenge * rlBreite * rlStaerke ) ) * cSPEZIFISCHES_GLASGEWICHT;
END_FUNCTION

(* ---- INC_UI.fn.st ---- *)
(* METADATA
{
	"v3Meta": {
		"objectGuid": "e071f047-ba29-40c0-bdd3-dce3563eb13b"
	}
}
*)
FUNCTION INC_UI : UINT
VAR_INPUT
  pui : REFERENCE TO UINT;
END_VAR
VAR
END_VAR

IF pui < 65536
THEN
  pui := pui + 1;
END_IF
END_FUNCTION

(* ---- INCI.fn.st ---- *)
(* METADATA
{
	"v3Meta": {
		"objectGuid": "47a21df2-edbb-49b0-932f-ef927933ed32"
	}
}
*)
FUNCTION INCI : INT
VAR_INPUT
  X : INT;
  N : INT;
END_VAR

(* Hinweis:
   - Funktion zum erhoehen der Eingangsvariablen X um 1. Sobald X den Wert N erreicht hat startet der Wert wieder bei 0.
*)
IF ( X >= N - 1 ) THEN
  INCI := 0;
ELSE
  INCI := X + 1;
END_IF;
END_FUNCTION

(* ---- INCW.fn.st ---- *)
(* METADATA
{
	"v3Meta": {
		"objectGuid": "c3800ee6-fccf-491b-bd53-b6c1155883a9"
	}
}
*)
FUNCTION INCW : WORD
VAR_INPUT
  X : WORD;
  N : WORD;
END_VAR

(* Hinweis:
   - Funktion zum erhoehen der Eingangsvariablen X um 1. Sobald X den Wert N erreicht hat startet der Wert wieder bei 0.
*)
IF ( X >= N - 1 ) THEN
  INCW := 0;
ELSE
  INCW := X + 1;
END_IF;
END_FUNCTION

(* ---- IsBetweenLReal.fn.st ---- *)
(* METADATA
{
	"v3Meta": {
		"objectGuid": "605f94de-cd86-43d0-95cd-83c44bc0f8dc"
	}
}
*)
FUNCTION IsBetweenLReal : BOOL
VAR_INPUT
  lriValue   : LREAL;
  lriBorder1 : LREAL;
  lriBorder2 : LREAL;
END_VAR
VAR
END_VAR

IsBetweenLReal := FALSE;

IF lriBorder1 < lriBorder2 THEN
  IsBetweenLReal := lriBorder1 <= lriValue
                    AND lriValue <= lriBorder2;
ELSE
  IsBetweenLReal := lriBorder2 <= lriValue
                    AND lriValue <= lriBorder1;
END_IF
END_FUNCTION

(* ---- IsBetweenWORD.fn.st ---- *)
(* METADATA
{
	"v3Meta": {
		"objectGuid": "640e1550-054d-48b5-a8dc-d9ce3f68325e"
	}
}
*)
FUNCTION IsBetweenWORD : BOOL
VAR_INPUT
  lwValue   : WORD;
  lwBorder1 : WORD;
  lwBorder2 : WORD;
END_VAR
VAR
END_VAR

IsBetweenWORD := FALSE;

IF lwBorder1 < lwBorder2 THEN
  IsBetweenWORD := lwBorder1 <= lwValue
                   AND lwValue <= lwBorder2;
ELSE
  IsBetweenWORD := lwBorder2 <= lwValue
                   AND lwValue <= lwBorder1;
END_IF
END_FUNCTION

(* ---- IsInRange.fn.st ---- *)
(* METADATA
{
	"v3Meta": {
		"objectGuid": "666a809c-7e52-4abd-9f01-34086fac7ebd"
	}
}
*)
FUNCTION IsInRange : BOOL
VAR_INPUT
  rlValue : REAL;
  rlTargetValue : REAL;
  rlThresshold : REAL;
END_VAR
VAR
END_VAR

IsInRange := ABS(rlValue - rlTargetValue) <= rlThresshold;
END_FUNCTION

(* ---- PruefungWertImIntervall.fn.st ---- *)
(* METADATA
{
	"v3Meta": {
		"objectGuid": "b7be4780-1c3e-4371-bb2a-cc9122a11be5"
	}
}
*)
FUNCTION PruefungWertImIntervall : BOOL
VAR_INPUT

  // WORD
  wpWert         : WORD;
  wpIntervallMin : WORD;
  wpIntervallMax : WORD;

END_VAR
VAR
END_VAR
//-------------------------------------------------------------------------------------------------
// LOGIK
//-------------------------------------------------------------------------------------------------
IF (  wpWert >= wpIntervallMin
     AND wpWert <= wpIntervallMax )
THEN
  PruefungWertImIntervall := TRUE;
ELSE
  PruefungWertImIntervall := FALSE;
END_IF
END_FUNCTION

(* ---- PruefungWertImIntervallAutomatikkreise.fn.st ---- *)
(* METADATA
{
	"v3Meta": {
		"objectGuid": "4fd29558-d6eb-46af-8028-798423b786a8"
	}
}
*)
FUNCTION PruefungWertImIntervallAutomatikkreise : BOOL
VAR_INPUT

  // WORD
  wpWert         : ARRAY[cERSTER_AUTOMATIKKREIS..cANZAHL_AUTOMATIKKREISE] OF Automatikkreis_EN;
  wpIntervallMin : WORD;
  wpIntervallMax : WORD;

END_VAR
VAR
  wlIndex : WORD;
END_VAR
//-------------------------------------------------------------------------------------------------
// LOGIK
//-------------------------------------------------------------------------------------------------
PruefungWertImIntervallAutomatikkreise := FALSE;

FOR wlIndex := cERSTER_AUTOMATIKKREIS TO cANZAHL_AUTOMATIKKREISE DO

  IF wpWert[wlIndex] = 0 THEN
    RETURN;
  END_IF

  IF (  wpWert[wlIndex] >= wpIntervallMin
       AND wpWert[wlIndex] <= wpIntervallMax )
  THEN
    PruefungWertImIntervallAutomatikkreise := TRUE;
  ELSE
    PruefungWertImIntervallAutomatikkreise := FALSE;
    RETURN;
  END_IF

END_FOR
END_FUNCTION

(* ---- RemoveETX.fn.st ---- *)
(* METADATA
{
	"v3Meta": {
		"objectGuid": "6a30dc93-6cfb-42ec-8e94-53fcaf08507e"
	}
}
*)
FUNCTION RemoveETX : ARRAY [0..3] OF DWORD
VAR_INPUT
  SheetID : ARRAY [0..3] OF DWORD;
END_VAR
VAR
  i, dwIn, dwOut, sh : INT;
  b : BYTE;
  tmp : DWORD;
END_VAR
FOR i := 0 TO 3 DO RemoveETX[i] := DWORD#0; END_FOR;

FOR i := 0 TO 15 DO
  dwIn := i / 4; sh := (i MOD 4) * 8;

  tmp := SHR(SheetID[dwIn], sh);     // byte runter schieben
  tmp := tmp MOD DWORD#256;          // entspricht AND 16#FF
  b := DWORD_TO_BYTE(tmp);

  IF b = BYTE#16#03 THEN b := BYTE#0; END_IF;

  dwOut := i / 4; sh := (i MOD 4) * 8;
  RemoveETX[dwOut] := RemoveETX[dwOut] + SHL(BYTE_TO_DWORD(b), sh);  // + statt OR
END_FOR;
END_FUNCTION

(* ---- ScheibenQuittierung.fn.st ---- *)
(* METADATA
{
	"v3Meta": {
		"objectGuid": "e5781056-5434-4b12-a4a2-e1c1e4aeb816"
	}
}
*)
FUNCTION ScheibenQuittierung : BOOL
VAR_INPUT

  // WORD
  wpQuellstation : WORD;
  wpZielStation  : WORD;
  wpQuellwand    : WORD := 1;
  wpZielwand     : WORD := 1;
  wpAuftragsTyp  : WORD := 0;

  // DWORD
  dwpWartezeit   : DWORD := 0;

END_VAR

VAR

  // BOOLEAN
  blResult : BOOL := FALSE;

END_VAR
//-------------------------------------------------------------------------------------------------
// FUNKTION: QUITTIEREN DER SCHEIBE
//-------------------------------------------------------------------------------------------------

wSps2MmiZielStation  := wpZielStation;
wSps2MmiQuellStation := wpQuellstation;
wSps2MmiZielWand     := wpZielwand;
wSps2MmiQuellWand    := wpQuellwand;
dwSps2MmiWartezeit   := dwpWartezeit;
wSPS2MMIAuftragstyp  := wpAuftragsTyp;

MsgToMmi(auftragsnr_w := SB0_SPS_QUIT_SHEET_ORDER );

ScheibenQuittierung := TRUE;
END_FUNCTION

(* ---- SendShuttlePosition.fn.st ---- *)
(* METADATA
{
	"v3Meta": {
		"objectGuid": "61256a4f-f80b-4fab-9669-5735e5c0be34"
	}
}
*)
FUNCTION SendShuttlePosition : BOOL
VAR_INPUT
END_VAR
VAR
  wlNummer : WORD;
  wlSlot   : WORD;
END_VAR
VAR CONSTANT
  cANZAHL_SLOTS_TELEGRAMM : WORD := 12; // Positionen die SB0_SPS_SORTIERUNGSHUTTLEPOS transportiert
END_VAR

//########################################## Changelog ################################################
//
//  2017-11-26 KV - Erstellt
//     => Function to send the current actual position of shuttle
//
//########################################## Changelog ################################################

(* Hinweis:
   - Die Position steht im MMI-Telegramm an einer festen Stelle (Slot), die Reihenfolge ist fest:
     1. Shuttles, 2. Transfershuttles, 3. Stationen die ein Shuttle sind [bStationIstShuttle]
   - Jede MK belegt einen Slot, auch wenn sie deaktiviert ist
   - Was nicht mehr ins Telegramm passt, wird nicht gesendet
*)
FOR wlSlot := 0 TO cANZAHL_SLOTS_TELEGRAMM - 1 DO
  rSps2MmiShuttlePosition[wlSlot] := 0.0;
END_FOR

wlSlot := 0;

// SHUTTLE
FOR wlNummer := cERSTES_SHUTTLE TO cLETZTES_SHUTTLE DO
  IF wlSlot < cANZAHL_SLOTS_TELEGRAMM THEN
    rSps2MmiShuttlePosition[wlSlot] := starrShuttleBasisParameter[wlNummer].rAktuellePositionQuerfahrt;
    wlSlot := wlSlot + 1;
  END_IF
END_FOR

// TRANSFERSHUTTLE
FOR wlNummer := cERSTES_TRANSFERSHUTTLE TO cLETZTES_TRANSFERSHUTTLE DO
  IF wlSlot < cANZAHL_SLOTS_TELEGRAMM THEN
    rSps2MmiShuttlePosition[wlSlot] := starrTransferShuttleBasisParameter[wlNummer].rAktuellePositionQuerfahrt;
    wlSlot := wlSlot + 1;
  END_IF
END_FOR

// STATIONEN die ein Shuttle sind
FOR wlNummer := cERSTE_STATION TO cLETZTE_STATION DO
  IF starrStationBasisParameter[wlNummer].stMKs.stSchnittstellendaten.bStationIstShuttle THEN
    IF wlSlot < cANZAHL_SLOTS_TELEGRAMM THEN
      rSps2MmiShuttlePosition[wlSlot] := starrStationBasisParameter[wlNummer].rAktuellePositionQuerfahrt;
      wlSlot := wlSlot + 1;
    END_IF
  END_IF
END_FOR

MsgToMmi(auftragsnr_w := SB0_SPS_SORTIERUNGSHUTTLEPOS);

SendShuttlePosition := TRUE;
END_FUNCTION

(* ---- setFreigabeKomponenten.fn.st ---- *)
(* METADATA
{
	"v3Meta": {
		"objectGuid": "691bf0f6-0a88-4d0a-9736-fcf4e429c02d"
	}
}
*)
FUNCTION setFreigabeKomponenten : BOOL
VAR_INPUT
  StationData : REFERENCE TO StationBasisParameter_ST;
END_VAR
VAR
  blSKAuswerten : BOOL; // Station hat gueltige MK, ist aktiv und hat mindestens einen SK konfiguriert
END_VAR
// Setzt alle Freigaben der Station (stFreigabe):
// - bAlles: NotHalt OK und ALLE Sicherheitskreise der Station geschlossen
// - bX    : NotHalt OK und alle SKs geschlossen, die Komponente X abschalten
//           (SK ohne Teilabschaltung schaltet alles ab, SK mit Teilabschaltung nur die markierten Komponenten)
// - Ohne konfigurierten SK (oder Station deaktiviert / keine MK): nur NotHalt
// - bgSicherheitstechnikBruecken setzt alle Freigaben

blSKAuswerten := checkSafetyCircuitsConfigured(StationData);

StationData.stFreigabe.bAlles           := ( NotHalt.bpNotHaltOK AND ( NOT blSKAuswerten OR_ELSE checkSafetyCircuitsClosed(StationData, eSKKomponente_Alles) ) )           OR bgSicherheitstechnikBruecken;
StationData.stFreigabe.bGlastransport   := ( NotHalt.bpNotHaltOK AND ( NOT blSKAuswerten OR_ELSE checkSafetyCircuitsClosed(StationData, eSKKomponente_Glastransport) ) )   OR bgSicherheitstechnikBruecken;
StationData.stFreigabe.bGeblaese        := ( NotHalt.bpNotHaltOK AND ( NOT blSKAuswerten OR_ELSE checkSafetyCircuitsClosed(StationData, eSKKomponente_Geblaese) ) )        OR bgSicherheitstechnikBruecken;
StationData.stFreigabe.bDrehen          := ( NotHalt.bpNotHaltOK AND ( NOT blSKAuswerten OR_ELSE checkSafetyCircuitsClosed(StationData, eSKKomponente_Drehen) ) )          OR bgSicherheitstechnikBruecken;
StationData.stFreigabe.bKippen          := ( NotHalt.bpNotHaltOK AND ( NOT blSKAuswerten OR_ELSE checkSafetyCircuitsClosed(StationData, eSKKomponente_Kippen) ) )          OR bgSicherheitstechnikBruecken;
StationData.stFreigabe.bQuerfahrt       := ( NotHalt.bpNotHaltOK AND ( NOT blSKAuswerten OR_ELSE checkSafetyCircuitsClosed(StationData, eSKKomponente_Querfahrt) ) )       OR bgSicherheitstechnikBruecken;
StationData.stFreigabe.bPneumatik       := ( NotHalt.bpNotHaltOK AND ( NOT blSKAuswerten OR_ELSE checkSafetyCircuitsClosed(StationData, eSKKomponente_Pneumatik) ) )       OR bgSicherheitstechnikBruecken;
StationData.stFreigabe.bGreifer         := ( NotHalt.bpNotHaltOK AND ( NOT blSKAuswerten OR_ELSE checkSafetyCircuitsClosed(StationData, eSKKomponente_Greifer) ) )         OR bgSicherheitstechnikBruecken;
StationData.stFreigabe.bWandverstellung := ( NotHalt.bpNotHaltOK AND ( NOT blSKAuswerten OR_ELSE checkSafetyCircuitsClosed(StationData, eSKKomponente_Wandverstellung) ) ) OR bgSicherheitstechnikBruecken;
StationData.stFreigabe.bMessachse       := ( NotHalt.bpNotHaltOK AND ( NOT blSKAuswerten OR_ELSE checkSafetyCircuitsClosed(StationData, eSKKomponente_Messachse) ) )       OR bgSicherheitstechnikBruecken;

setFreigabeKomponenten := StationData.stFreigabe.bAlles;
END_FUNCTION

(* ---- SetWatchIO.fn.st ---- *)
(* METADATA
{
	"v3Meta": {
		"objectGuid": "35aa6819-3357-423e-91ac-0c94eb5a5c7a"
	}
}
*)
FUNCTION SetWatchIO : Bool
VAR_INPUT
  in_Word   : WORD;
  in_Number : WORD;
END_VAR
VAR
  wIndex    : WORD;
END_VAR

FOR wIndex := 0 TO 15 DO
  WatchIo(((in_Word AND (SHL(1, wIndex))) <> 0), (in_Number - 1) + (wIndex + 1));
END_FOR;

//ChangedBits := in_Word XOR old_Word;
//
//IF ChangedBits <> 0 THEN
//
//    FOR i := 0 TO 15 DO
//        IF (ChangedBits AND (SHL(1 , i))) <> 0 THEN
//            WatchIo(((in_Word AND ( SHL(1, i))) <> 0), (in_Number -1) +(i+1) );
//        END_IF;
//    END_FOR;
//  old_Word := in_Word; // alten Wert speichern
//END_IF;
END_FUNCTION

(* ---- StationHatShuttleNachbar.fn.st ---- *)
(* METADATA
{
	"v3Meta": {
		"objectGuid": "1fe72243-ca8e-4332-9b86-e73fbf76fe1f"
	}
}
*)
FUNCTION StationHatShuttleNachbar : BOOL
VAR_IN_OUT CONSTANT
  stpBasis : StationBasisParameter_ST;
END_VAR
VAR
  wlNachbar : WORD;
  stlNachbar : REFERENCE TO StationBasisParameter_ST;
END_VAR

(* Hinweis:
   - TRUE, wenn ein konfigurierter Ein- oder Austransport-Partner der Station ein Shuttle ist
     [MK stSchnittstellendaten.bStationIstShuttle, kann auch bei einer Station gesetzt sein]
   - Im Systemcheck kann eine Scheibe dann zum Teil noch auf dem Shuttle liegen,
     eine abweichende Belegung ist deshalb nur ein Hinweis und kein Fehler
*)
StationHatShuttleNachbar := FALSE;

IF NOT __ISVALIDREF( stpBasis.stMKs ) THEN
  RETURN;
END_IF

FOR wlNachbar := cERSTES_SHUTTLE TO cLETZTE_FREMDANLAGE_EINLAUF DO

  IF    ( stpBasis.stMKs.stSchnittstellendaten.aEintransporte.Station[wlNachbar] <> TransportRichtung_EN.Default )
     OR ( stpBasis.stMKs.stSchnittstellendaten.aAustransporte.Station[wlNachbar] <> TransportRichtung_EN.Default )
  THEN
    stlNachbar REF= getBasis( wlNachbar );

    IF     __ISVALIDREF( stlNachbar )
       AND_THEN __ISVALIDREF( stlNachbar.stMKs )
       AND_THEN stlNachbar.stMKs.stSchnittstellendaten.bStationIstShuttle
    THEN
      StationHatShuttleNachbar := TRUE;
      RETURN;
    END_IF
  END_IF

END_FOR
END_FUNCTION

(* ---- StationInAutomatikkreis.fn.st ---- *)
(* METADATA
{
	"v3Meta": {
		"objectGuid": "a9180b59-ead2-48cb-98e6-a6809a238554"
	}
}
*)
FUNCTION StationInAutomatikkreis : BOOL
VAR_INPUT
  awpArray : ARRAY[cERSTER_AUTOMATIKKREIS..cANZAHL_AUTOMATIKKREISE] OF Automatikkreis_EN;
  wpValueToFind : WORD;
END_VAR
VAR
  INDEX : WORD;
END_VAR

StationInAutomatikkreis := FALSE;

FOR INDEX := cERSTER_AUTOMATIKKREIS TO cANZAHL_AUTOMATIKKREISE DO

  IF awpArray[INDEX] = wpValueToFind THEN
    StationInAutomatikkreis := TRUE;
    RETURN;
  END_IF

END_FOR
END_FUNCTION

(* ---- StationInSicherheitskreis.fn.st ---- *)
(* METADATA
{
	"v3Meta": {
		"objectGuid": "28064981-b681-426a-a86e-e794fcbf1911"
	}
}
*)
FUNCTION StationInSicherheitskreis : BOOL
VAR_INPUT
  awpArray : ARRAY[0..cANZAHL_SICHERHEITSKREISE] OF Sicherheitskreis_EN;
  wpValueToFind : WORD;
END_VAR
VAR
  INDEX : WORD;
END_VAR

StationInSicherheitskreis := FALSE;

FOR INDEX := 0 TO cANZAHL_SICHERHEITSKREISE DO

  IF awpArray[INDEX] = wpValueToFind THEN
    StationInSicherheitskreis := TRUE;
    RETURN;
  END_IF

END_FOR
END_FUNCTION

(* ---- TransferShuttleBetriebsstopAktiv.fn.st ---- *)
(* METADATA
{
	"v3Meta": {
		"objectGuid": "00eb9e03-2e2c-414f-a437-451e0f99c47c"
	}
}
*)
FUNCTION TransferShuttleBetriebsstopAktiv : BOOL
VAR_INPUT
  eAutomatikkreis : Automatikkreis_EN;
END_VAR
VAR
  wlIndex : WORD;
END_VAR

TransferShuttleBetriebsstopAktiv := FALSE;

FOR wlIndex := cERSTES_TRANSFERSHUTTLE TO cLETZTES_TRANSFERSHUTTLE DO

  IF NOT starrTransfershuttleBasisParameter[wlIndex].stMKs.bDeaktivieren THEN

    IF StationInAutomatikkreis(starrTransfershuttleBasisParameter[wlIndex].stMKs.eaAutomatikkreis, eAutomatikkreis) THEN
      IF aTransfershuttles[wlIndex].bpAnforderungBetriebsstopp THEN
        TransferShuttleBetriebsstopAktiv := TRUE;
        RETURN;
      END_IF
    END_IF
  END_IF
END_FOR
END_FUNCTION

(* ---- WegZumScheibenTrennenBestimmen.fn.st ---- *)
(* METADATA
{
	"v3Meta": {
		"objectGuid": "975fc77d-048f-43ed-b0dc-a9d95a26ef34"
	}
}
*)
FUNCTION WegZumScheibenTrennenBestimmen : REAL
VAR_INPUT

  // REAL
  rpAuftragsLaenge       : REAL := REAL#0; // [mm]
  rpRampe                : REAL := 1000.0; // [mm/s^2] Verzoegerungsrampe  => Werte muessen umgerechnet werden in [m/s^2]
  rpGeschwindigkeit      : REAL := 1000;   // [m/s]   Sollgeschwindigkeit => Werte muessen umgerechnet werden in [m/s]
  rpTrennGeschwindigkeit : REAL := 500;    // [m/s]   Geschwindigkeit mit der die Beladung aufgetrennt werden soll => Werte muessen umgerechnet werden in [m/s]

END_VAR
VAR

  // REAL
  rlBerechneteTrennStrecke         : REAL := REAL#0;
  rlBerechneteVerzoegerungsStrecke : REAL := REAL#0;
  rlValidierungWert                : REAL := REAL#0;
  rlRueckgabeWert                  : REAL := REAL#0;

END_VAR
VAR CONSTANT

  // REAL
  cVALIDIERUNG_NULL             : REAL := REAL#0;
  cVALIDIERUNGSWERT             : REAL := 100.0;
  cDEFAULT_RAMPE                : REAL := 1000.0;
  cDEFAULT_GESCHWINDIGKEIT      : REAL := 1000.0;
  cDEFAULT_TRENNGESCHWINDIGKEIT : REAL := 500.0;

  // WORD
  cMILLIMETER_ZU_METER_FAKTOR   : WORD := 1000;

END_VAR
// Info:
//   - Es wird mittels uebergebener Daten ein Weg berechnet ab wann der Antrieb verzoegern muss, um
//     eine Stationsbeladung sauber aufzutrennen.

//-------------------------------------------------------------------------------------------------
// FUNKTION: ERMITTELN EINER STRECKE ZUM TRENNEN EINER STATIONSBELADUNG
//-------------------------------------------------------------------------------------------------
(* Hinweis:
   - Auftragslaenge muss angegeben werden
*)
IF ( rpAuftragsLaenge <= 0 ) THEN
  WegZumScheibenTrennenBestimmen := REAL#0;
  RETURN;
END_IF

(* Hinweis:
   - Sicherstellen das keine 0 Rampen bzw. keine 0 Geschwindigkeit angegeben wurde
     => Fuellen mit default Werten (Division durch null Verhindern)
*)
IF ( ABS(rpRampe) <= cVALIDIERUNG_NULL ) THEN
  rpRampe := cDEFAULT_RAMPE;
END_IF

IF ( ABS(rpGeschwindigkeit) <= cVALIDIERUNG_NULL ) THEN
  rpGeschwindigkeit := cDEFAULT_GESCHWINDIGKEIT;
END_IF

IF ( ABS(rpTrennGeschwindigkeit) <= cVALIDIERUNG_NULL ) THEN
  rpTrennGeschwindigkeit := cDEFAULT_TRENNGESCHWINDIGKEIT;
END_IF

(* Hinweis:
   - Werte in die passende pysikalische Einheit umwandeln
     => Rampe von mm/s^2 zu m/s^2
     => Geschwindigkeit von mm/s zu m/s
     => Laenge von mm zu m
*)
rpRampe                 := ABS( rpRampe / cMILLIMETER_ZU_METER_FAKTOR );
rpGeschwindigkeit       := ABS( rpGeschwindigkeit / cMILLIMETER_ZU_METER_FAKTOR );
rpTrennGeschwindigkeit  := ABS( rpTrennGeschwindigkeit / cMILLIMETER_ZU_METER_FAKTOR );
rpAuftragsLaenge        := ABS( rpAuftragsLaenge / cMILLIMETER_ZU_METER_FAKTOR );

(* Hinweis:
   - Strecke berechnen die benoetigt wird, um von der Soll- Geschwindigkeit auf die reduzierte
     Trenn- Geschwindigkeit zu kommen
      => s =  v^2 - v0^2 / 2*a
*)
rlBerechneteTrennStrecke := LREAL_TO_REAL(ABS((EXPT(rpGeschwindigkeit,2) - EXPT(rpTrennGeschwindigkeit,2)) / ( 2 * rpRampe )));

(* Hinweis:
   - Strecke berechnen die gebraucht wird, wenn aus maximaler (Soll-) Geschwindigkeit abgebremst wird
     => S = v^2 / (2*a)
*)
rlBerechneteVerzoegerungsStrecke := LREAL_TO_REAL((EXPT(rpGeschwindigkeit,2) ) / ( 2 * rpRampe ));

(* Hinweis:
   - Strecken summieren
*)
rlValidierungWert :=  ( ( rpAuftragsLaenge - ( rlBerechneteVerzoegerungsStrecke + rlBerechneteTrennStrecke) ) * cMILLIMETER_ZU_METER_FAKTOR );

IF ( rlValidierungWert <= cVALIDIERUNGSWERT ) THEN
  rlRueckgabeWert := REAL#0;

ELSE
  rlRueckgabeWert := rlValidierungWert;

END_IF

WegZumScheibenTrennenBestimmen := rlRueckgabeWert;
END_FUNCTION
